(* IEC 61131-3 sources: sis-interlock-demo/tests/POUs/Suites/FB_VoteEval_Test, 7 files *)

(* ---- ArchHelpersChannelsAndRequired.method.decl.st ---- *)
// F_VoteArchChannels и F_VoteArchRequired: N и M по таблице 5.1, 0 для None, ForcedTrip и вне перечисления
METHOD PRIVATE ArchHelpersChannelsAndRequired
VAR
    uBad : U_SisEnumInt;   // значение вне перечисления
END_VAR

(* ---- ArchNoneTripsReportsNone.method.decl.st ---- *)
// Схема None и ForcedTrip как заданная схема: срабатывание, действующая схема None, без деградации,
// счётчики 0 — даже если все каналы в норме
METHOD PRIVATE ArchNoneTripsReportsNone
VAR
    aeCh  : ARRAY[1..GVL_Const.SIS_VOTE_CH_MAX] OF E_ChannelState;   // состояния каналов
    stRes : ST_VoteResult;                                           // результат
END_VAR

(* ---- ChannelsBeyondNIgnored.method.decl.st ---- *)
// Каналы с номером больше N не голосуют: 1oo1 с требованием на каналах 2 и 3 — нет срабатывания
METHOD PRIVATE ChannelsBeyondNIgnored
VAR
    aeCh  : ARRAY[1..GVL_Const.SIS_VOTE_CH_MAX] OF E_ChannelState;   // состояния каналов
    stRes : ST_VoteResult;                                           // результат
END_VAR

(* ---- CountersReportStates.method.decl.st ---- *)
// Счётчики D, F, B, H равны числу каналов в каждом состоянии
METHOD PRIVATE CountersReportStates
VAR
    aeCh  : ARRAY[1..GVL_Const.SIS_VOTE_CH_MAX] OF E_ChannelState;   // состояния каналов
    stRes : ST_VoteResult;                                           // результат
END_VAR

(* ---- NotUsedInsideNCountsInvalid.method.decl.st ---- *)
// NotUsed и значение вне перечисления внутри N считаются недостоверными каналами (безопасная сторона)
METHOD PRIVATE NotUsedInsideNCountsInvalid
VAR
    aeCh  : ARRAY[1..GVL_Const.SIS_VOTE_CH_MAX] OF E_ChannelState;   // состояния каналов
    stRes : ST_VoteResult;                                           // результат
    uBad  : U_SisEnumInt;                                            // значение вне перечисления
END_VAR

(* ---- PolicyOutOfEnumTripsNone.method.decl.st ---- *)
// Политика вне перечисления (7): срабатывание, схема None, счётчики 0
METHOD PRIVATE PolicyOutOfEnumTripsNone
VAR
    aeCh  : ARRAY[1..GVL_Const.SIS_VOTE_CH_MAX] OF E_ChannelState;   // состояния каналов
    stRes : ST_VoteResult;                                           // результат
    uBad  : U_SisEnumInt;                                            // значение вне перечисления
END_VAR

(* ---- TwoOfThreeTripsOnSecondDemand.method.decl.st ---- *)
// 2oo3 без деградации: один канал Demand — нет срабатывания, два — срабатывание; схема 2oo3
METHOD PRIVATE TwoOfThreeTripsOnSecondDemand
VAR
    aeCh  : ARRAY[1..GVL_Const.SIS_VOTE_CH_MAX] OF E_ChannelState;   // состояния каналов
    stRes : ST_VoteResult;                                           // результат
END_VAR
